// TIA Portal V21 export
// export: Created 2026-11-10T07:35:00.8181146Z, ExportSetting WithDefaults, DisplayName Totally Integrated Automation Portal, DisplayVersion V21 Update 3, DisplayName STEP 7 Professional, DisplayVersion V21 Update 3, DisplayName STEP 7 Safety, DisplayVersion V21, DisplayName Tech WebApplication, DisplayVersion V21, DisplayName WinCC Basic/Comfort/Advanced, DisplayVersion V21 Update 3, DisplayName WinCC Unified, DisplayVersion V21 Update 3
FUNCTION_BLOCK "FB_Lad_ex005"   // FB5, LAD
{ S7_Optimized_Access := 'TRUE' }
VERSION : 0.1
// stored: AutoNumber true, IsIECCheckEnabled false, IsRetainMemResEnabled false, MemoryReserve 100, SetENOAutomatically false, UDAEnableTagReadback false
   VAR_INPUT
      v_in1 : DTL;
      v_in2 : DTL;
      v_out : Time;
   END_VAR
BEGIN

REGION Network 1: T_DIFF - Time difference
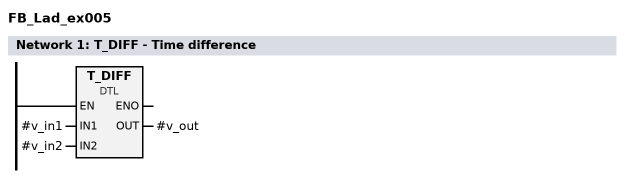
   RUNG wire#powerrail
      { S7_Templates := "[date_type := DTL, time_type := Time]" } T_DIFF(IN1 := #v_in1, IN2 := #v_in2, OUT => #v_out)
   END_RUNG
   // the same network as SCL:
   T_DIFF(IN1 := #v_in1, IN2 := #v_in2, OUT => #v_out);
END_REGION
END_FUNCTION_BLOCK
